// TIA Portal V21 export
DATA_BLOCK "IDB_SclCalls"   // DB18
// stored: InstanceOfName FB_SclCalls, InstanceOfType FB
"FB_SclCalls"
   // VAR_INPUT
   //    Enable : Bool;
   //    Mode : Int;
   //    Delta : Real;
   // END_VAR
   // VAR_OUTPUT
   //    Average : Real;
   //    Scaled : Real;
   //    CallsOk : Bool;
   // END_VAR
   // VAR_IN_OUT
   //    TimerBlock : "FB_SclTimers";
   //    Values : Array[0..9] of Real;
   // END_VAR
   // VAR
   //    Sections { S7_SetPoint := 'True'} : "FB_SclSections";
   //    Total : LReal;
   //    Rounded : DInt;
   //    ResultText : String;
   //    Magnitude : Real;
   //    ConvertedWord : Word;
   //    IntValue : Int;
   //    ShortValue : SInt;
   //    NarrowValue : Int;
   // END_VAR
BEGIN
END_DATA_BLOCK
